(* PLC project g_hvac_fan_delay_clean, Anonymous Benchmark Suite 1.0 *)
(* stored: creationDateTime 2026-07-09T00:00:00 *)

PROGRAM g_hvac_fan_delay_clean
  VAR_INPUT
    heat_call : BOOL;
    cool_call : BOOL;
    enable : BOOL;
    maint : BOOL;
  END_VAR
  VAR_OUTPUT
    heat : BOOL;
    cool : BOOL;
    fan : BOOL;
  END_VAR

(* LD diagram, written out as Structured Text *)
heat := NOT cool_call AND heat_call AND enable;
cool := cool_call AND enable;
fan := enable;
END_PROGRAM

CONFIGURATION Config0
  RESOURCE Res0 ON PLC
    TASK tcyclic(INTERVAL := T#10ms, PRIORITY := 0);
    PROGRAM inst0 WITH tcyclic : g_hvac_fan_delay_clean;
  END_RESOURCE
END_CONFIGURATION
